PROGRAM main
  VAR
    B1 AT %IX0.0     : BOOL; (* sensor de cajas *)
    KM1 AT %QX0.0    : BOOL; (* banda (bobina 00001 para la PC) *)
    CAJAS AT %MW0    : INT; (* holding 40001: cajas contadas *)
    P_MARCHA AT %MW1 : INT; (* holding 40002: pulsador remoto MARCHA *)
    P_PARO AT %MW2   : INT; (* holding 40003: pulsador remoto PARO *)
    P_CERO AT %MW3   : INT; (* holding 40004: pulsador remoto contador a cero *)
    F_CAJA           : R_TRIG;
    CAJA             : BOOL; (* flanco de B1 *)
  END_VAR
  VAR  (* added by the conversion: wires and edge detectors of the diagram *)
    _ADD7_OUT : INT;
    _SEL4_OUT : INT;
    _NE14_OUT : BOOL;
    _OR12_OUT : BOOL;
    _EQ17_OUT : BOOL;
    _AND11_OUT : BOOL;
    _NE22_OUT : BOOL;
    _SEL21_OUT : INT;
    _NE29_OUT : BOOL;
    _SEL28_OUT : INT;
  END_VAR

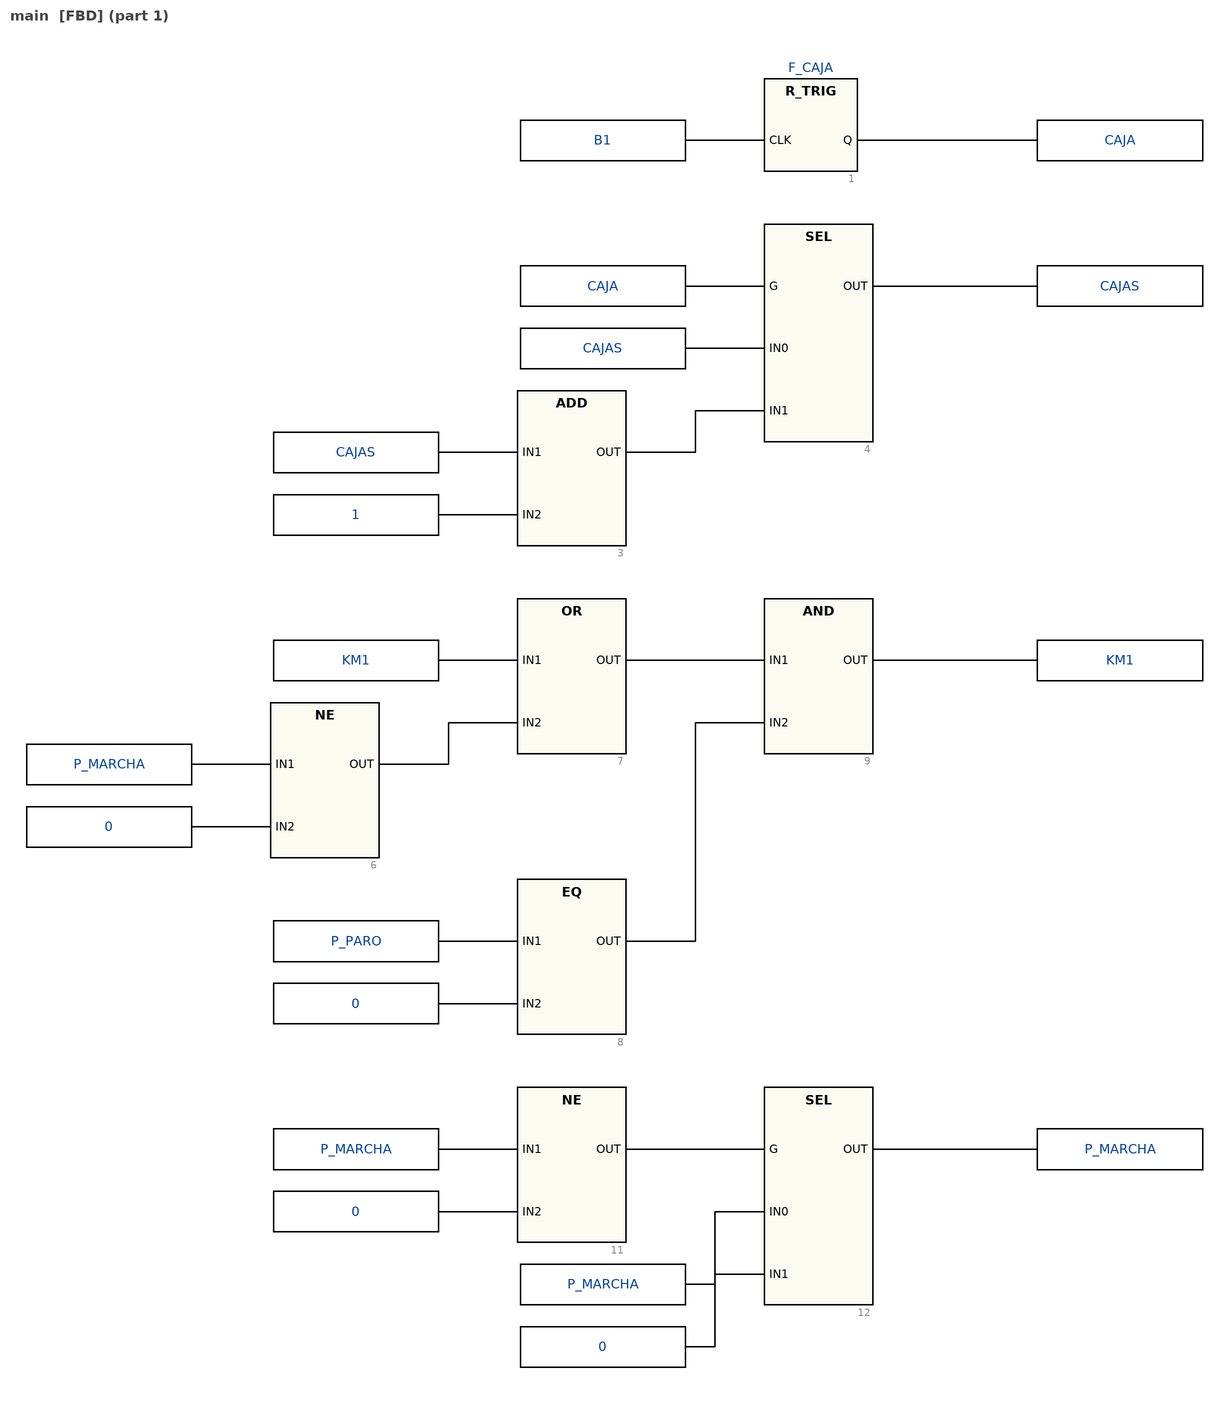
(* FBD diagram, written out as Structured Text *)
F_CAJA(CLK := B1);
CAJA := F_CAJA.Q;
_ADD7_OUT := CAJAS + 1;
_SEL4_OUT := SEL(CAJA, CAJAS, _ADD7_OUT);
CAJAS := _SEL4_OUT;
_NE14_OUT := P_MARCHA <> 0;
_OR12_OUT := KM1 OR _NE14_OUT;
_EQ17_OUT := P_PARO = 0;
_AND11_OUT := _OR12_OUT AND _EQ17_OUT;
KM1 := _AND11_OUT;
_NE22_OUT := P_MARCHA <> 0;
_SEL21_OUT := SEL(_NE22_OUT, P_MARCHA, 0);
P_MARCHA := _SEL21_OUT;
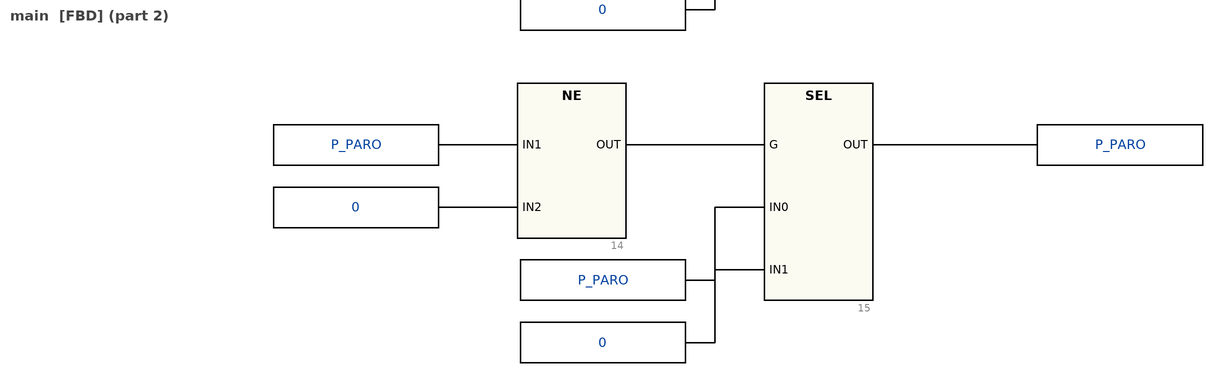
_NE29_OUT := P_PARO <> 0;
_SEL28_OUT := SEL(_NE29_OUT, P_PARO, 0);
P_PARO := _SEL28_OUT;
END_PROGRAM
